PROGRAM MAIN
VAR
END_VAR

GVL_IO.xLaserEnable := NOT GVL_IO.xNotHalt_Betaetigt;

END_PROGRAM

(* stored: Version 1.1.0.1
   POU MAIN: Id {44c38e53-312d-458f-a823-461371afcb42}, SpecialFunc None *)
